(* IEC 61131-3 sources: plc-st-coding-agent/progress/evidence/full_r8_20261110b/native_evidence/codex_minimax-m27/public-medium-07/0, 1 file *)

(* ---- candidate.st ---- *)
FUNCTION_BLOCK FB
VAR_INPUT
    OCCUPANCY_DETECTED    : BOOL;
    ENERGY_SAVING_MODE    : BOOL;
    HVAC_MODE_SELECTOR    : INT;
END_VAR
VAR_OUTPUT
    SUPPLY_FAN_RUN        : BOOL := FALSE;
    TEMP_SETPOINT_ADJUST  : INT  := 0;
END_VAR
VAR
    OccupancyCounter      : INT := 0;
END_VAR

// Temperature setpoint adjustment (initialized at power-up)
IF HVAC_MODE_SELECTOR = 0 THEN
    IF OCCUPANCY_DETECTED THEN
        TEMP_SETPOINT_ADJUST := 0;
    ELSIF ENERGY_SAVING_MODE THEN
        TEMP_SETPOINT_ADJUST := 3;
    ELSE
        TEMP_SETPOINT_ADJUST := 2;
    END_IF
ELSIF HVAC_MODE_SELECTOR = 1 THEN
    IF OCCUPANCY_DETECTED THEN
        TEMP_SETPOINT_ADJUST := 0;
    ELSE
        TEMP_SETPOINT_ADJUST := 1;
    END_IF
ELSIF HVAC_MODE_SELECTOR = 2 THEN
    IF OCCUPANCY_DETECTED THEN
        TEMP_SETPOINT_ADJUST := 0;
    ELSE
        TEMP_SETPOINT_ADJUST := 4;
    END_IF
ELSE
    TEMP_SETPOINT_ADJUST := 4;
END_IF

IF TEMP_SETPOINT_ADJUST > 4 THEN
    TEMP_SETPOINT_ADJUST := 4;
ELSIF TEMP_SETPOINT_ADJUST < -4 THEN
    TEMP_SETPOINT_ADJUST := -4;
END_IF;

// Supply fan delay control: 30-scan delay, level-reset
IF OCCUPANCY_DETECTED AND HVAC_MODE_SELECTOR <> 3 THEN
    IF OccupancyCounter < 30 THEN
        OccupancyCounter := OccupancyCounter + 1;
    END_IF;
    IF OccupancyCounter >= 30 THEN
        SUPPLY_FAN_RUN := TRUE;
    ELSE
        SUPPLY_FAN_RUN := FALSE;
    END_IF;
ELSE
    OccupancyCounter := 0;
    SUPPLY_FAN_RUN := FALSE;
END_IF;

END_FUNCTION_BLOCK
